// TIA Portal V19 export
FUNCTION "Alarms" : Void   // FC2, LAD
{ S7_Optimized_Access := 'TRUE' }
// stored: SetENOAutomatically false
BEGIN

REGION Network 1: Alarm
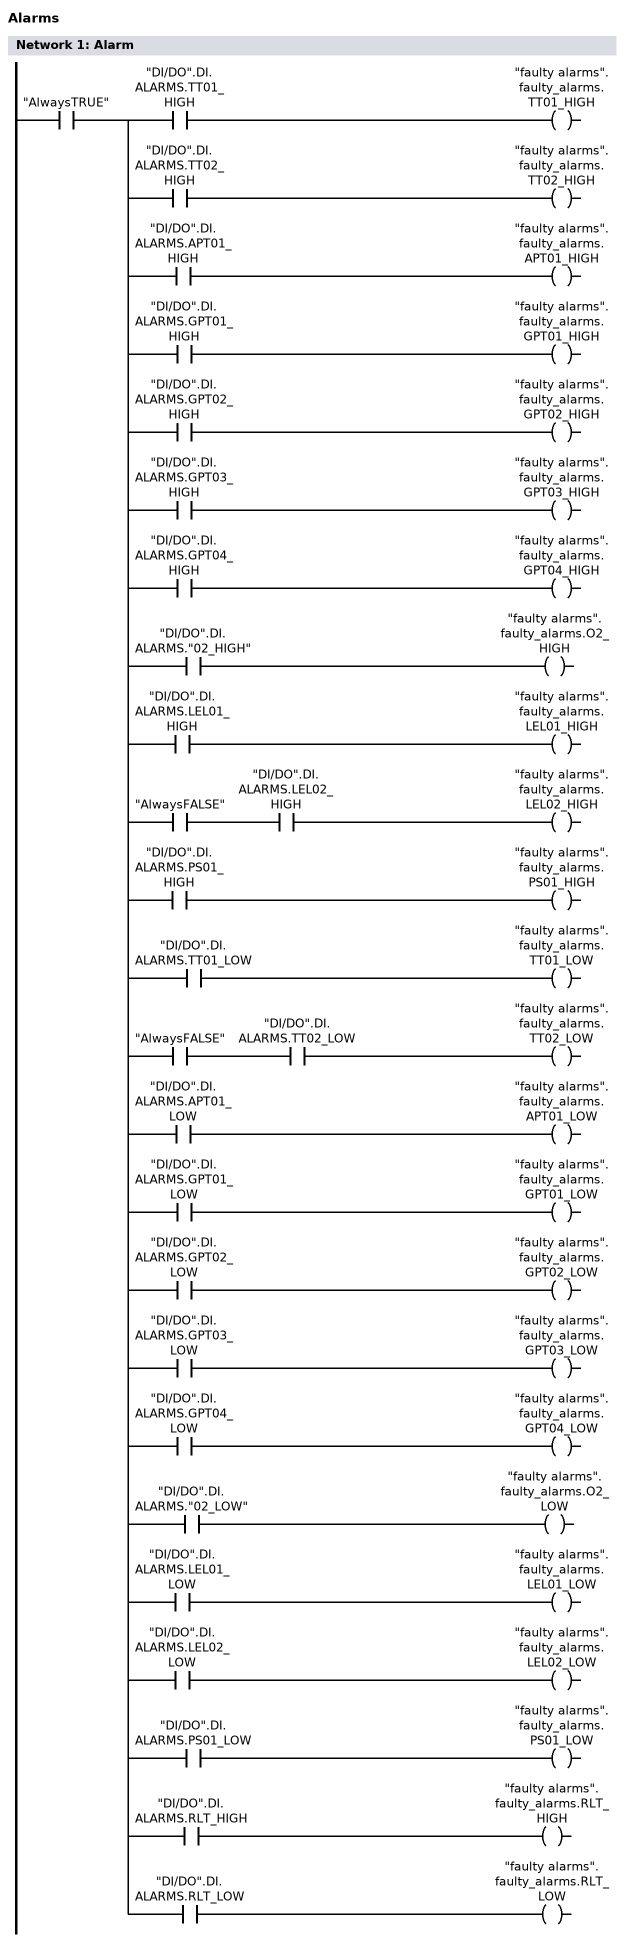
   RUNG wire#powerrail
      Contact( "AlwaysTRUE" )
      wire#w1
      Contact( "DI/DO".DI.ALARMS.TT01_HIGH )
      Coil( "faulty alarms".faulty_alarms.TT01_HIGH )
   END_RUNG
   RUNG wire#w1
      Contact( "DI/DO".DI.ALARMS.TT02_HIGH )
      Coil( "faulty alarms".faulty_alarms.TT02_HIGH )
   END_RUNG
   RUNG wire#w1
      Contact( "DI/DO".DI.ALARMS.APT01_HIGH )
      Coil( "faulty alarms".faulty_alarms.APT01_HIGH )
   END_RUNG
   RUNG wire#w1
      Contact( "DI/DO".DI.ALARMS.GPT01_HIGH )
      Coil( "faulty alarms".faulty_alarms.GPT01_HIGH )
   END_RUNG
   RUNG wire#w1
      Contact( "DI/DO".DI.ALARMS.GPT02_HIGH )
      Coil( "faulty alarms".faulty_alarms.GPT02_HIGH )
   END_RUNG
   RUNG wire#w1
      Contact( "DI/DO".DI.ALARMS.GPT03_HIGH )
      Coil( "faulty alarms".faulty_alarms.GPT03_HIGH )
   END_RUNG
   RUNG wire#w1
      Contact( "DI/DO".DI.ALARMS.GPT04_HIGH )
      Coil( "faulty alarms".faulty_alarms.GPT04_HIGH )
   END_RUNG
   RUNG wire#w1
      Contact( "DI/DO".DI.ALARMS."02_HIGH" )
      Coil( "faulty alarms".faulty_alarms.O2_HIGH )
   END_RUNG
   RUNG wire#w1
      Contact( "DI/DO".DI.ALARMS.LEL01_HIGH )
      Coil( "faulty alarms".faulty_alarms.LEL01_HIGH )
   END_RUNG
   RUNG wire#w1
      Contact( "AlwaysFALSE" )
      Contact( "DI/DO".DI.ALARMS.LEL02_HIGH )
      Coil( "faulty alarms".faulty_alarms.LEL02_HIGH )
   END_RUNG
   RUNG wire#w1
      Contact( "DI/DO".DI.ALARMS.PS01_HIGH )
      Coil( "faulty alarms".faulty_alarms.PS01_HIGH )
   END_RUNG
   RUNG wire#w1
      Contact( "DI/DO".DI.ALARMS.TT01_LOW )
      Coil( "faulty alarms".faulty_alarms.TT01_LOW )
   END_RUNG
   RUNG wire#w1
      Contact( "AlwaysFALSE" )
      Contact( "DI/DO".DI.ALARMS.TT02_LOW )
      Coil( "faulty alarms".faulty_alarms.TT02_LOW )
   END_RUNG
   RUNG wire#w1
      Contact( "DI/DO".DI.ALARMS.APT01_LOW )
      Coil( "faulty alarms".faulty_alarms.APT01_LOW )
   END_RUNG
   RUNG wire#w1
      Contact( "DI/DO".DI.ALARMS.GPT01_LOW )
      Coil( "faulty alarms".faulty_alarms.GPT01_LOW )
   END_RUNG
   RUNG wire#w1
      Contact( "DI/DO".DI.ALARMS.GPT02_LOW )
      Coil( "faulty alarms".faulty_alarms.GPT02_LOW )
   END_RUNG
   RUNG wire#w1
      Contact( "DI/DO".DI.ALARMS.GPT03_LOW )
      Coil( "faulty alarms".faulty_alarms.GPT03_LOW )
   END_RUNG
   RUNG wire#w1
      Contact( "DI/DO".DI.ALARMS.GPT04_LOW )
      Coil( "faulty alarms".faulty_alarms.GPT04_LOW )
   END_RUNG
   RUNG wire#w1
      Contact( "DI/DO".DI.ALARMS."02_LOW" )
      Coil( "faulty alarms".faulty_alarms.O2_LOW )
   END_RUNG
   RUNG wire#w1
      Contact( "DI/DO".DI.ALARMS.LEL01_LOW )
      Coil( "faulty alarms".faulty_alarms.LEL01_LOW )
   END_RUNG
   RUNG wire#w1
      Contact( "DI/DO".DI.ALARMS.LEL02_LOW )
      Coil( "faulty alarms".faulty_alarms.LEL02_LOW )
   END_RUNG
   RUNG wire#w1
      Contact( "DI/DO".DI.ALARMS.PS01_LOW )
      Coil( "faulty alarms".faulty_alarms.PS01_LOW )
   END_RUNG
   RUNG wire#w1
      Contact( "DI/DO".DI.ALARMS.RLT_HIGH )
      Coil( "faulty alarms".faulty_alarms.RLT_HIGH )
   END_RUNG
   RUNG wire#w1
      Contact( "DI/DO".DI.ALARMS.RLT_LOW )
      Coil( "faulty alarms".faulty_alarms.RLT_LOW )
   END_RUNG
   // the same network as SCL:
   "faulty alarms".faulty_alarms.TT01_HIGH := "AlwaysTRUE" AND "DI/DO".DI.ALARMS.TT01_HIGH;
   "faulty alarms".faulty_alarms.TT02_HIGH := "AlwaysTRUE" AND "DI/DO".DI.ALARMS.TT02_HIGH;
   "faulty alarms".faulty_alarms.APT01_HIGH := "AlwaysTRUE" AND "DI/DO".DI.ALARMS.APT01_HIGH;
   "faulty alarms".faulty_alarms.GPT01_HIGH := "AlwaysTRUE" AND "DI/DO".DI.ALARMS.GPT01_HIGH;
   "faulty alarms".faulty_alarms.GPT02_HIGH := "AlwaysTRUE" AND "DI/DO".DI.ALARMS.GPT02_HIGH;
   "faulty alarms".faulty_alarms.GPT03_HIGH := "AlwaysTRUE" AND "DI/DO".DI.ALARMS.GPT03_HIGH;
   "faulty alarms".faulty_alarms.GPT04_HIGH := "AlwaysTRUE" AND "DI/DO".DI.ALARMS.GPT04_HIGH;
   "faulty alarms".faulty_alarms.O2_HIGH := "AlwaysTRUE" AND "DI/DO".DI.ALARMS."02_HIGH";
   "faulty alarms".faulty_alarms.LEL01_HIGH := "AlwaysTRUE" AND "DI/DO".DI.ALARMS.LEL01_HIGH;
   "faulty alarms".faulty_alarms.LEL02_HIGH := "AlwaysTRUE" AND "AlwaysFALSE" AND "DI/DO".DI.ALARMS.LEL02_HIGH;
   "faulty alarms".faulty_alarms.PS01_HIGH := "AlwaysTRUE" AND "DI/DO".DI.ALARMS.PS01_HIGH;
   "faulty alarms".faulty_alarms.TT01_LOW := "AlwaysTRUE" AND "DI/DO".DI.ALARMS.TT01_LOW;
   "faulty alarms".faulty_alarms.TT02_LOW := "AlwaysTRUE" AND "AlwaysFALSE" AND "DI/DO".DI.ALARMS.TT02_LOW;
   "faulty alarms".faulty_alarms.APT01_LOW := "AlwaysTRUE" AND "DI/DO".DI.ALARMS.APT01_LOW;
   "faulty alarms".faulty_alarms.GPT01_LOW := "AlwaysTRUE" AND "DI/DO".DI.ALARMS.GPT01_LOW;
   "faulty alarms".faulty_alarms.GPT02_LOW := "AlwaysTRUE" AND "DI/DO".DI.ALARMS.GPT02_LOW;
   "faulty alarms".faulty_alarms.GPT03_LOW := "AlwaysTRUE" AND "DI/DO".DI.ALARMS.GPT03_LOW;
   "faulty alarms".faulty_alarms.GPT04_LOW := "AlwaysTRUE" AND "DI/DO".DI.ALARMS.GPT04_LOW;
   "faulty alarms".faulty_alarms.O2_LOW := "AlwaysTRUE" AND "DI/DO".DI.ALARMS."02_LOW";
   "faulty alarms".faulty_alarms.LEL01_LOW := "AlwaysTRUE" AND "DI/DO".DI.ALARMS.LEL01_LOW;
   "faulty alarms".faulty_alarms.LEL02_LOW := "AlwaysTRUE" AND "DI/DO".DI.ALARMS.LEL02_LOW;
   "faulty alarms".faulty_alarms.PS01_LOW := "AlwaysTRUE" AND "DI/DO".DI.ALARMS.PS01_LOW;
   "faulty alarms".faulty_alarms.RLT_HIGH := "AlwaysTRUE" AND "DI/DO".DI.ALARMS.RLT_HIGH;
   "faulty alarms".faulty_alarms.RLT_LOW := "AlwaysTRUE" AND "DI/DO".DI.ALARMS.RLT_LOW;
END_REGION
END_FUNCTION
